FUNCTION F_MoveToAxisRef : ST_PLCTOSTOEBER
VAR_IN_OUT
	Axis							:ST_AXIS_REF;				(* The AXIS_REF data type  is an interface between the PLC and the NC and contains axis information *)
END_VAR
VAR_INPUT
	stTerminalState				:ST_TerminalState;
	stStoeberToPlc				:ST_STOEBERTOPLC;
END_VAR
VAR
END_VAR

(* Set terminal parameters *)
Axis.sAdsAddr:= F_CreateAmsNetId(stTerminalState.stAdsAddr.netId);
Axis.unSlaveAddr:= stTerminalState.stAdsAddr.port;

(* Copy the actual values from the inverter to the axis reference *)
Axis.stNcToPlc.stBaseDevice.bEnabled := stStoeberToPlc.byE200DeviceStatusByte.0;			(* The drive is ready for operation. *)
Axis.stNcToPlc.stBaseDevice.bError := stStoeberToPlc.byE200DeviceStatusByte.1;				(* The drive state is fault. *)
Axis.stNcToPlc.stBaseDevice.bGroupError := stStoeberToPlc.unI200PosiStatusWord.2;			(* Group error: Maximum following error *)
Axis.stNcToPlc.stBaseDevice.bQuickStop := stStoeberToPlc.byE200DeviceStatusByte.2;			(* Quick stop is queued/is being executed. *)
Axis.stNcToPlc.stBaseDevice.bAxisActive := stStoeberToPlc.byE200DeviceStatusByte.5;			(* Axis is active. *)
Axis.stNcToPlc.stBaseDevice.bToggleBit := stStoeberToPlc.byE200DeviceStatusByte.7;			(* Handshake bit. *)

Axis.stNcToPlc.stBaseDevice.stCommandPositioning.bConstantVelocity := stStoeberToPlc.unI200PosiStatusWord.4;			(* Constant speed reached. *)
Axis.stNcToPlc.stBaseDevice.stCommandPositioning.bHomed := stStoeberToPlc.unI200PosiStatusWord.6;					(* Axis is referenced. *)
Axis.stNcToPlc.stBaseDevice.stCommandPositioning.bPositionReached := stStoeberToPlc.unI200PosiStatusWord.5;			(* Window around target position reached for the first time. *)
Axis.stNcToPlc.stBaseDevice.stCommandPositioning.bPositionWinReached := stStoeberToPlc.byI201MotionStatusByte.5;		(* Actual position is located in the position window. *)
Axis.stNcToPlc.stBaseDevice.stCommandPositioning.bNotMoving := NOT stStoeberToPlc.byE200DeviceStatusByte.0           	(* Control enabled *) 			(* Axis is logically stationary. *)
               										     			      OR NOT stStoeberToPlc.byE200DeviceStatusByte.5     	(* An axis is active. *)
               										     			      OR stStoeberToPlc.unI200PosiStatusWord.7;                          (* Axis standstill *)
Axis.stNcToPlc.stBaseDevice.stCommandPositioning.bDenied := stStoeberToPlc.unI200PosiStatusWord.1;					(* Indicates that the command denied .*)
Axis.stNcToPlc.stBaseDevice.stCommandPositioning.bCoupled := (stStoeberToPlc.byI201MotionStatusByte AND 16#0F) = 5;	(* Axis coupling state *)
Axis.stNcToPlc.stBaseDevice.stCommandPositioning.dnActPosition := stStoeberToPlc.dnI203CurrentPosition;				(* Value of current (actual) position *)
Axis.stNcToPlc.stBaseDevice.stCommandPositioning.dnActVelocity := stStoeberToPlc.dnI88Speed;						(* Value of current (actual) velocity *)
Axis.stNcToPlc.stBaseDevice.stCommandPositioning.nActEngineTorque := stStoeberToPlc.nE90MMotor;					(* Indication of the current motor torque in Nm *)

Axis.stNcToPlc.stBaseDevice.stCommandPositioning.bLimitMaxExceeded := NOT Axis.stPlcToNc.stBaseDevice.bFeedEnablePlus;		(* Position limit switch maximum is exceeded *)
Axis.stNcToPlc.stBaseDevice.stCommandPositioning.bLimitMinExceeded := NOT Axis.stPlcToNc.stBaseDevice.bFeedEnableMinus;		(* Position limit switch minimum is exceeded *)

Axis.stNcToPlc.stBaseDevice.stCommandPositioning.byPLCOpenState := stStoeberToPlc.byI201MotionStatusByte AND 2#00001111;				(* Supplies information on the reaction of the axis during operation on a fieldbus. *)
Axis.stNcToPlc.stBaseDevice.stCommandPositioning.bPLCOpenStandstill := stStoeberToPlc.unI200PosiStatusWord.7;							(* PLCopen state Standstill. *)
Axis.stNcToPlc.stBaseDevice.stCommandPositioning.bPLCOpenCmdAborted :=  stStoeberToPlc.unI200PosiStatusWord.3;						(* Positioning command denied/aborted. TRUE means that the last positioning job was aborted. *)
Axis.stNcToPlc.stBaseDevice.stCommandPositioning.bPLCOpenCmdDone := stStoeberToPlc.byI201MotionStatusByte.4;							(* TRUE means that the command was executed successfully. *)
Axis.stNcToPlc.stBaseDevice.stCommandPositioning.byPLCOpenErrorCode := stStoeberToPlc.byI90ErrorCode;									(* When the PLCOpen state is ErrorStop. *)

Axis.stNcToPlc.stBaseDevice.stFastRefereneValue.bStandstill := stStoeberToPlc.nD200SpeedReferenceValueStatusWord.0;						(* Standstill. *)
Axis.stNcToPlc.stBaseDevice.stFastRefereneValue.bVeloReached := stStoeberToPlc.nD200SpeedReferenceValueStatusWord.1;					(* Reference value reached *)
Axis.stNcToPlc.stBaseDevice.stFastRefereneValue.nMotorSpeed := stStoeberToPlc.nE100MMotor;											(* Current motor speed *)

(* Copy the setpoint values from the axis reference to the inverter *)
F_MoveToAxisRef.byA180DeviceControlByte.0 := Axis.stPlcToNc.stBaseDevice.bEnable;				(* Enable controller *)
F_MoveToAxisRef.byA180DeviceControlByte.1 := Axis.stPlcToNc.stBaseDevice.bFaultReset;				(* Acknowledgment for faults of the device state machine. *)
F_MoveToAxisRef.byA180DeviceControlByte.2 := Axis.stPlcToNc.stBaseDevice.bQuickStop;				(* Brakes the motor *)
F_MoveToAxisRef.wI210PosiControlWord.1 := Axis.stPlcToNc.stBaseDevice.bFeedEnablePlus;			(* Feed enable plus *)
F_MoveToAxisRef.wI210PosiControlWord.2 := Axis.stPlcToNc.stBaseDevice.bFeedEnableMinus;			(* Feed enable minus *)
F_MoveToAxisRef.wI210PosiControlWord.3 :=  Axis.stPlcToNc.stBaseDevice.bHomingSensor;			(* Referencing cam signal or homing sensor *)
F_MoveToAxisRef.byA180DeviceControlByte.7 :=  Axis.stPlcToNc.stBaseDevice.bToggleBit;				(* Handshake bit. *)
F_MoveToAxisRef.nC230TorqueLimit	 := Axis.stPlcToNc.stBaseDevice.nTorqueLimit;						(* Value of torque limit (absolute value) *)

F_MoveToAxisRef.nI230Override := Axis.stPlcToNc.stBaseDevice.stCommandPositioning.nOverride;							(* Value of override 16384 = 100 %. *)
F_MoveToAxisRef.nI215VeloFaktor := Axis.stPlcToNc.stBaseDevice.stCommandPositioning.nVeloFactor;						(* Value of the velocity 16384 = 100 %. *)
F_MoveToAxisRef.usnI216AccFaktor := Axis.stPlcToNc.stBaseDevice.stCommandPositioning.usnAccFactor;					(* Value of the acceleration (always positive) 255 = 100% *)
F_MoveToAxisRef.usnI217DccFaktor := Axis.stPlcToNc.stBaseDevice.stCommandPositioning.usnDccFaktor	;				(* Value of the deceleration (always positive) 255 = 100% *)
F_MoveToAxisRef.dnI213TargetPosition := Axis.stPlcToNc.stBaseDevice.stCommandPositioning.dnTargetPosition;				(* Value of target position *)
F_MoveToAxisRef.dnI34ReferencePosition := Axis.stPlcToNc.stBaseDevice.stCommandPositioning.dnReferencePosition;			(* Value which is loaded as the actual position in the reference point.  *)
F_MoveToAxisRef.wI210PosiControlWord.4 := Axis.stPlcToNc.stBaseDevice.stCommandPositioning.bTipEnable;				(* Activates tipping mode. *)
F_MoveToAxisRef.wI210PosiControlWord.5 := Axis.stPlcToNc.stBaseDevice.stCommandPositioning.bTipPlus;					(* Tip mode in positive direction. *)
F_MoveToAxisRef.wI210PosiControlWord.6 := Axis.stPlcToNc.stBaseDevice.stCommandPositioning.bTipMinus;					(* Tip mode in negative direction. *)
F_MoveToAxisRef.byI211MotionCommandByte := Axis.stPlcToNc.stBaseDevice.stCommandPositioning.byPLCOpenCmd;			(* Global parameter for specification of the command to be executed via fieldbus. *)
F_MoveToAxisRef.wI210PosiControlWord.0 := Axis.stPlcToNc.stBaseDevice.stCommandPositioning.bPLCOpenCmdExe;			(* With a rising edge, the command in Motion Command is executed. *)

F_MoveToAxisRef.nD230NReferenceValueRelative := Axis.stPlcToNc.stBaseDevice.stFastRefereneValue.nSpeed;				(* Relative speed reference value *)

END_FUNCTION

(* stored: Version 1.1.0.1, ProductVersion 3.1.4024.15
   POU F_MoveToAxisRef: Id {1ba4e7e8-1871-46fd-a8f7-08c63d7efe44}, SpecialFunc None *)
